// Mitsubishi GX Works2 project: 261012_타이머실습_타이머추가응용3   PLC: Q03UDV

PROGRAM MAIN
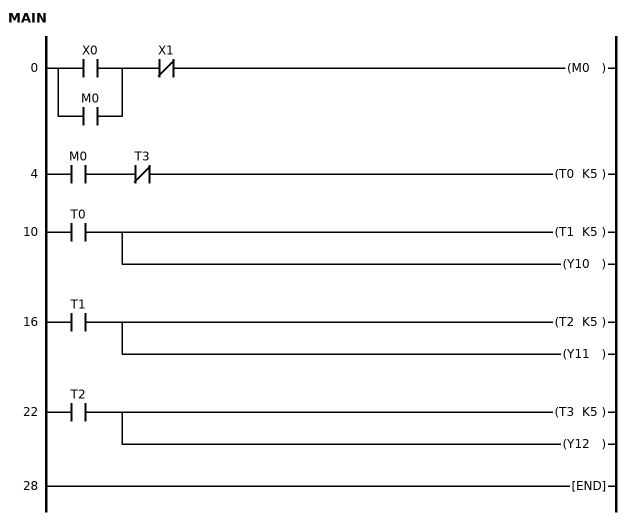
0     LD      X0
      OR      M0
      ANI     X1
      OUT     M0
4     LD      M0
      ANI     T3
      OUT     T0 K5
10    LD      T0
      OUT     T1 K5
      OUT     Y10
16    LD      T1
      OUT     T2 K5
      OUT     Y11
22    LD      T2
      OUT     T3 K5
      OUT     Y12
28    END
END_PROGRAM
